FUNCTION F_MGR_TO_OPC (* OPC-UA-Endpunkt aus MGR_ID: 192.168.1.12:61499 -> opc.tcp://192.168.1.12:4840 *)
  (* Standard: 61499-1; Description: Copyright (c) 2026 Meisterschulen am Ostbahnhof This program and the accompanying materials are made available under the terms of the Eclipse Public License 2.0 which is available at https://www.eclipse.org/legal/epl-2.0/ SPDX-License-Identifier: EPL-2.0 *)
  (* Version 1.0, 2026-10-17, Franz Höpfinger, Meisterschulen am Ostbahnhof, initial implementation *)
  PACKAGE MyLib_OPC;
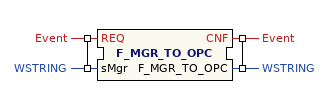
  EVENT_INPUT
    REQ WITH sMgr;
  END_EVENT
  EVENT_OUTPUT
    CNF WITH F_MGR_TO_OPC;
  END_EVENT
  VAR_INPUT
    sMgr : WSTRING; (* MGR_ID der Station, z.B. logiBUS::stations::Computers::C_12 *)
  END_VAR
  VAR_OUTPUT
    F_MGR_TO_OPC : WSTRING;
  END_VAR
  BODY IN ST:
PACKAGE MyLib_OPC;

(* OPC-UA-Endpunkt aus MGR_ID: 192.168.1.12:61499 -> opc.tcp://192.168.1.12:4840 *)
FUNCTION F_MGR_TO_OPC : WSTRING

VAR_INPUT
	sMgr : WSTRING; // MGR_ID der Station, z.B. logiBUS::stations::Computers::C_12
END_VAR

F_MGR_TO_OPC := CONCAT("opc.tcp://", LEFT(sMgr, FIND(sMgr, ":")), "4840");

END_FUNCTION
  END_BODY
END_FUNCTION
